// TIA Portal V21 export
// export: Created 2026-10-23T20:43:33.5103753Z, ExportSetting WithDefaults, DisplayName Totally Integrated Automation Portal, DisplayVersion V21 Update 1, DisplayName SINAMICS Startdrive Advanced, DisplayVersion V21 HF2, DisplayName SINAMICS Startdrive G110M, G120, G120C, G120D, G120P, G115D, DisplayVersion V21 HF2, DisplayName SINAMICS Startdrive G130, G150, S120, S150, G200, G220, S200, S210, S220, Innomotics MVD, DisplayVersion V21 HF2, DisplayName STEP 7 Professional, DisplayVersion V21 Update 1, DisplayName STEP 7 Safety, DisplayVersion V21, DisplayName Tech WebApplication, DisplayVersion V21, DisplayName WinCC Basic/Comfort/Advanced, DisplayVersion V21 Update 1, DisplayName WinCC Unified, DisplayVersion V21 Update 1
FUNCTION_BLOCK "FB_AnaForCounter"   // FB20, SCL
TITLE = Analyzer: FOR counter modified
{ S7_Optimized_Access := 'TRUE' }
VERSION : 0.1
// Rule C26h: the FOR counter Index is changed inside the loop through the reference IndexRef (TIA refuses a direct or InOut change)
// stored: AutoNumber true, IsIECCheckEnabled false, IsRetainMemResEnabled false, MemoryReserve 100, SetENOAutomatically false, UDAEnableTagReadback false
   VAR_INPUT
      Limit : Int;   // Stop when the total exceeds this
   END_VAR
   VAR_OUTPUT
      Total : Int;   // Sum of the indices
   END_VAR
   VAR
      Index : Int;   // Loop counter
   END_VAR
   VAR_TEMP
      IndexRef : REF_TO Int;   // Reference to the loop counter
   END_VAR
BEGIN

       #Total := 0;
       #IndexRef := REF(#Index);
       FOR #Index := 0 TO 10 DO
           #Total := #Total + #Index;
           IF #Total > #Limit THEN
               #IndexRef^ := 10;
           END_IF;
       END_FOR;
END_FUNCTION_BLOCK
